Universal Robots URScript: T011_zai-org_GLM-4.7-FP8_edit_perf_rep1.urscript

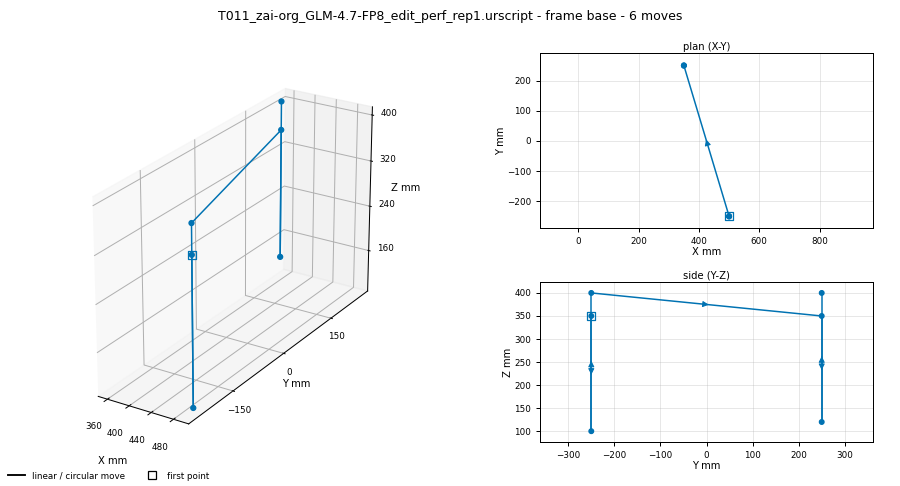
[picture p0: tool path of T011_zai-org_GLM-4.7-FP8_edit_perf_rep1.urscript in frame base, 6 of 8 moves have a stored position in this frame; points joined in program order, loops and branches not executed]
# Task: T011 — Dual-zone pick-place — hybrid mode (OPTIMIZED)
# Generated by ENFIELD IR→URScript Translator
# Operating mode: hybrid | Max TCP speed: 0.300 m/s
# Robot: ur5e
#
# WARNING: This is auto-generated code for SIMULATION ONLY.
# Do NOT deploy to a physical robot without safety review.

def task_T011():
  # [0] E-Stop verify
  # E-Stop safety check (hardware-enforced on UR controller)
  if (get_digital_in(0) == True):
    popup("E-Stop active — aborting program.", error=True)
    halt
  end

  # [1] Home
  # Increased joint velocity and acceleration for faster repositioning
  movej([0.0000, -1.5708, 1.5708, -1.5708, -1.5708, 0.0000], a=2.0000, v=1.2000)

  # [2] Above storage bin
  # Maximized linear speed to limit, increased acceleration
  movel(p[0.500000, -0.250000, 0.350000, 0.0000, 3.1416, 0.0000], a=1.2000, v=0.3000, r=0.0200)

  # [3] Descend to pick
  # Increased speed significantly for faster cycle, kept slightly below max for precision
  movel(p[0.500000, -0.250000, 0.100000, 0.0000, 3.1416, 0.0000], a=1.0000, v=0.2500)

  # [4] Gripper CLOSE
  # Gripper CLOSE (force=50 N)
  set_digital_out(0, True)

  # [5] Grip settle
  # Reduced sleep time to minimize cycle delay
  sleep(0.1000)

  # [6] Lift from bin
  # Maximized speed, increased blend radius for smoother transition
  movel(p[0.500000, -0.250000, 0.400000, 0.0000, 3.1416, 0.0000], a=1.2000, v=0.3000, r=0.0300)

  # [7] Transit to handoff zone
  # Maximized speed and acceleration, increased blend radius
  movel(p[0.350000, 0.250000, 0.350000, 0.0000, 3.1416, 0.0000], a=1.5000, v=0.3000, r=0.0400)

  # [8] Place at handoff
  # Increased speed for placement
  movel(p[0.350000, 0.250000, 0.120000, 0.0000, 3.1416, 0.0000], a=0.8000, v=0.2000)

  # [9] Gripper OPEN
  # Gripper OPEN
  set_digital_out(0, False)

  # [10] Release
  # Reduced sleep time
  sleep(0.1000)

  # [11] Retract
  # Maximized speed
  movel(p[0.350000, 0.250000, 0.400000, 0.0000, 3.1416, 0.0000], a=1.2000, v=0.3000, r=0.0200)

  # [12] Return home
  # Increased joint velocity and acceleration
  movej([0.0000, -1.5708, 1.5708, -1.5708, -1.5708, 0.0000], a=2.0000, v=1.2000)

end

# Entry point
task_T011()
